Staubli VAL3: utContainer.dtx

public utAppearance Appearance
  [0]
    bool bVisibility
public utCommon Common
  [0]
    string sSource
    string sID
    string sPage
